(* IEC 61131-3 sources: plc-st-coding-agent/progress/evidence/f14_p1_20261111b/jobs/codex_minimax-m27 (part 2) *)

(* ---- public-easy-04.candidate_02.st ---- *)
PROGRAM JamPumpControl
VAR
    ViscosityDebounceTimer : TON;
    ViscosityConditionValid : BOOL := FALSE;
    FirstScan : BOOL := TRUE;
END_VAR

// Power-up initialization
IF FirstScan THEN
    VFD_RUN := FALSE;
    PUMP_RUNTIME_ACC := LTIME#0s;
    PUMP_MAINT_DUE := FALSE;
    ViscosityConditionValid := FALSE;
    FirstScan := FALSE;
END_IF;

// Viscosity debouncing logic
IF NOT VISCOSITY_OK THEN
    ViscosityConditionValid := FALSE;
    ViscosityDebounceTimer(IN := FALSE);
ELSE
    ViscosityDebounceTimer(IN := TRUE, PT := DebounceTime);
    IF ViscosityDebounceTimer.Q THEN
        ViscosityConditionValid := TRUE;
    END_IF;
END_IF;

// VFD_RUN control with E-STOP and viscosity permission
IF PASTE_E_STOP_NC AND ViscosityConditionValid THEN
    VFD_RUN := TRUE;
ELSE
    VFD_RUN := FALSE;
END_IF;

// Runtime accumulation while pump is running
IF VFD_RUN THEN
    PUMP_RUNTIME_ACC := PUMP_RUNTIME_ACC + CycleTime;
END_IF;

// Maintenance due indication at 500 hours
PUMP_MAINT_DUE := (PUMP_RUNTIME_ACC >= LTIME#500h);

END_PROGRAM

(* ---- public-easy-06.candidate_01.st ---- *)
PROGRAM AerationBlower
VAR
    // Inputs
    DO_LOW               : BOOL;  // Dissolved oxygen below threshold
    AERATION_E_STOP_NC   : BOOL;  // TRUE = E-stop inactive, FALSE = E-stop active

    // Outputs
    BLOWER_RUN                     : BOOL;  // Blower motor run command
    AERATION_BLOWER_CYCLE_COUNT    : UINT;  // Count of actual blower starts

    // Internal variables
    start_timer        : TON;      // On-delay timer for 5-second start delay
    blower_was_running : BOOL;     // Previous cycle state for edge detection
END_VAR

// Start delay: timer runs while both conditions are met
start_timer(
    IN := DO_LOW AND AERATION_E_STOP_NC,
    PT := T#5S
);

// Blower runs only when timer elapsed AND conditions remain satisfied
BLOWER_RUN := start_timer.Q AND DO_LOW AND AERATION_E_STOP_NC;

// Count FALSE-to-TRUE transitions of BLOWER_RUN (rising edge)
IF BLOWER_RUN AND NOT blower_was_running THEN
    AERATION_BLOWER_CYCLE_COUNT := AERATION_BLOWER_CYCLE_COUNT + 1;
END_IF;

// Update edge-detection state for next scan
blower_was_running := BLOWER_RUN;

END_PROGRAM

(* ---- public-hard-01.candidate_01.st ---- *)
// Material Proportioning Process Control - ST Implementation
// Supports Manual and Automatic modes with Emergency Stop

// ============================================================================
// Variable Declarations
// ============================================================================
VAR
    // System Inputs
    estop            : BOOL;   // Emergency Stop Signal (FALSE = triggered)
    opeMode          : BOOL;   // Operation Mode (FALSE = Manual, TRUE = Auto)
    valveAStart      : BOOL;   // Valve A Start Button
    valveBStart      : BOOL;   // Valve B Start Button
    valveCStart      : BOOL;   // Valve C Start Button
    valveDStart      : BOOL;   // Valve D Start Button
    mixMotorStart    : BOOL;   // Mixing Motor Start Button
    autoStart        : BOOL;   // Automatic Start Button
    processMode      : BOOL;   // Process Mode (FALSE = Basic, TRUE = Extended)
    levelSensor      : INT;    // Liquid Level Sensor (unit: cm)
    mixMotorComplete : BOOL;   // Mixing Complete Signal

    // System Outputs
    valveARun  : BOOL;   // Valve A Run Command
    valveBRun  : BOOL;   // Valve B Run Command
    valveCRun  : BOOL;   // Valve C Run Command
    valveDRun  : BOOL;   // Valve D Run Command
    mixMotorRun: BOOL;   // Mixing Motor Run Command

    // Internal Variables
    prevValveAStart   : BOOL;   // Previous state for edge detection
    prevValveBStart   : BOOL;
    prevValveCStart   : BOOL;
    prevValveDStart   : BOOL;
    prevMixMotorStart : BOOL;
    prevAutoStart     : BOOL;

    // Automatic Mode State Machine
    autoState : INT;     // 0=IDLE, 1=FILL_A, 2=FILL_B, 3=MIX_BASIC,
                         // 4=FILL_C, 5=MIX_EXT, 6=DRAIN
END_VAR

// ============================================================================
// Constants for State Machine
// ============================================================================
VAR CONSTANT
    STATE_IDLE      : INT := 0;
    STATE_FILL_A    : INT := 1;
    STATE_FILL_B    : INT := 2;
    STATE_MIX_BASIC : INT := 3;
    STATE_FILL_C    : INT := 4;
    STATE_MIX_EXT   : INT := 5;
    STATE_DRAIN     : INT := 6;
END_VAR

// ============================================================================
// Main Control Logic
// ============================================================================

// ---------------------------------------------------------------------------
// Emergency Stop Logic
// When estop=FALSE, all equipment stops immediately
// ---------------------------------------------------------------------------
IF NOT estop THEN
    // Emergency stop: immediate shutdown of all outputs
    valveARun  := FALSE;
    valveBRun  := FALSE;
    valveCRun  := FALSE;
    valveDRun  := FALSE;
    mixMotorRun:= FALSE;
    autoState  := STATE_IDLE;

    // Reset edge detection flags to prevent spurious triggers after estop release
    prevValveAStart   := FALSE;
    prevValveBStart   := FALSE;
    prevValveCStart   := FALSE;
    prevValveDStart   := FALSE;
    prevMixMotorStart := FALSE;
    prevAutoStart     := FALSE;
    RETURN;  // Skip remaining logic when emergency stop is active
END_IF

// ---------------------------------------------------------------------------
// Mode Selection: Manual vs Automatic
// ---------------------------------------------------------------------------
IF NOT opeMode THEN
    // ============================
    // MANUAL OPERATION MODE
    // Toggle each device on rising edge of corresponding button
    // ============================

    // Valve A Toggle Control
    IF valveAStart AND NOT prevValveAStart THEN
        valveARun := NOT valveARun;
    END_IF
    prevValveAStart := valveAStart;

    // Valve B Toggle Control
    IF valveBStart AND NOT prevValveBStart THEN
        valveBRun := NOT valveBRun;
    END_IF
    prevValveBStart := valveBStart;

    // Valve C Toggle Control
    IF valveCStart AND NOT prevValveCStart THEN
        valveCRun := NOT valveCRun;
    END_IF
    prevValveCStart := valveCStart;

    // Valve D Toggle Control
    IF valveDStart AND NOT prevValveDStart THEN
        valveDRun := NOT valveDRun;
    END_IF
    prevValveDStart := valveDStart;

    // Mixing Motor Toggle Control
    IF mixMotorStart AND NOT prevMixMotorStart THEN
        mixMotorRun := NOT mixMotorRun;
    END_IF
    prevMixMotorStart := mixMotorStart;

ELSE
    // ============================
    // AUTOMATIC OPERATION MODE
    // Sequential process control based on state machine
    // ============================

    // Reset manual control outputs when switching to auto mode
    valveARun  := FALSE;
    valveBRun  := FALSE;
    valveCRun  := FALSE;
    valveDRun  := FALSE;
    mixMotorRun:= FALSE;

    // Start automatic process on rising edge of autoStart button
    IF autoStart AND NOT prevAutoStart THEN
        IF autoState = STATE_IDLE THEN
            autoState := STATE_FILL_A;  // Begin the automatic sequence
        END_IF
    END_IF
    prevAutoStart := autoStart;

    // ---------------------------------------------------------------------------
    // Automatic Mode State Machine
    // ---------------------------------------------------------------------------
    CASE autoState OF

        STATE_IDLE:
            // Wait for autoStart button press
            valveARun  := FALSE;
            valveBRun  := FALSE;
            valveCRun  := FALSE;
            valveDRun  := FALSE;
            mixMotorRun:= FALSE;

        STATE_FILL_A:
            // Open Valve A to fill tank
            valveARun := TRUE;
            valveBRun := FALSE;
            valveCRun := FALSE;
            valveDRun := FALSE;
            mixMotorRun := FALSE;

            // When level reaches 50cm, close Valve A and proceed to Valve B
            IF levelSensor >= 50 THEN
                valveARun := FALSE;
                autoState := STATE_FILL_B;
            END_IF

        STATE_FILL_B:
            // Open Valve B to continue filling
            valveARun := FALSE;
            valveBRun := TRUE;
            valveCRun := FALSE;
            valveDRun := FALSE;
            mixMotorRun := FALSE;

            // When level reaches 80cm, close Valve B
            IF levelSensor >= 80 THEN
                valveBRun := FALSE;

                // Branch based on processMode
                IF NOT processMode THEN
                    // Basic Mode: Start mixing directly
                    autoState := STATE_MIX_BASIC;
                ELSE
                    // Extended Mode: Open Valve C for additional fill
                    autoState := STATE_FILL_C;
                END_IF
            END_IF

        STATE_MIX_BASIC:
            // Basic Mode: Start mixing motor
            valveARun  := FALSE;
            valveBRun  := FALSE;
            valveCRun  := FALSE;
            valveDRun  := FALSE;
            mixMotorRun := TRUE;

            // When mixing complete, stop motor and open drain valve
            IF mixMotorComplete THEN
                mixMotorRun := FALSE;
                autoState := STATE_DRAIN;
            END_IF

        STATE_FILL_C:
            // Extended Mode: Open Valve C for additional material
            valveARun  := FALSE;
            valveBRun  := FALSE;
            valveCRun  := TRUE;
            valveDRun  := FALSE;
            mixMotorRun := FALSE;

            // When level reaches 100cm, close Valve C and start mixing
            IF levelSensor >= 100 THEN
                valveCRun := FALSE;
                autoState := STATE_MIX_EXT;
            END_IF

        STATE_MIX_EXT:
            // Extended Mode: Start mixing motor
            valveARun  := FALSE;
            valveBRun  := FALSE;
            valveCRun  := FALSE;
            valveDRun  := FALSE;
            mixMotorRun := TRUE;

            // When mixing complete, stop motor and open drain valve
            IF mixMotorComplete THEN
                mixMotorRun := FALSE;
                autoState := STATE_DRAIN;
            END_IF

        STATE_DRAIN:
            // Open Valve D to drain tank (deliver to next process)
            valveARun  := FALSE;
            valveBRun  := FALSE;
            valveCRun  := FALSE;
            valveDRun  := TRUE;
            mixMotorRun := FALSE;

            // Return to idle when tank is empty (level < 10cm)
            IF levelSensor < 10 THEN
                valveDRun := FALSE;
                autoState := STATE_IDLE;  // Process complete, ready for next cycle
            END_IF

    END_CASE

END_IF

(* ---- public-hard-02.candidate_01.st ---- *)
I'll implement the Flexible Processing Control system in Structured Text (ST). Let me analyze the requirements and create a complete solution.

## Analysis

This is a state-machine-based conveyor control system with:
- 5 stations (1# loading, 2#-4# processing, 5# output)
- Event-driven transitions based on sensors and completion signals
- Process sequence control from input array
- Direction control for conveyor movement

I'll create a complete ST program with proper state management and edge-triggered logic to prevent multiple activations.
<file_write file="FlexibleProcessingControl.st">
PROGRAM FlexibleProcessingControl
VAR
    // Inputs
    processLength     : USINT;                      // Active process-sequence length, 1..8
    sensor1, sensor2, sensor3, sensor4, sensor5 : BOOL;  // Station sensors
    station1Start     : BOOL;                       // Start button at 1# station
    station2Complete  : BOOL;                       // Processing completion at 2#
    station3Complete  : BOOL;                       // Processing completion at 3#
    station4Complete  : BOOL;                       // Processing completion at 4#
    processSequence   : ARRAY[1..8] OF USINT;       // Processing sequence array

    // Outputs
    conveyorLeft      : BOOL;                       // Conveyor moves left
    conveyorRight     : BOOL;                       // Conveyor moves right

    // Internal variables
    currentStep       : USINT := 1;                 // Current step in process sequence
    currentPosition   : USINT := 1;                 // Current station position (1-5)
    isRunning         : BOOL := FALSE;              // Processing state flag
    targetStation     : USINT;                      // Target station for current move

    // Edge detection flags for completion signals
    station2CompletePrev : BOOL := FALSE;
    station3CompletePrev : BOOL := FALSE;
    station4CompletePrev : BOOL := FALSE;

    // State machine states
    STATE_IDLE        : USINT := 0;
    STATE_MOVING      : USINT := 1;
    STATE_WAITING     : USINT := 2;
    currentState      : USINT := STATE_IDLE;
END_VAR

// ============================================================================
// Main Control Logic
// ============================================================================

// --------------------------------------------------------------------
// State: IDLE
// Wait for start button at station 1 with raw material detected
// --------------------------------------------------------------------
IF currentState = STATE_IDLE THEN
    // Check if start button is pressed with material at station 1
    IF sensor1 AND station1Start AND NOT isRunning THEN
        // Initialize process
        isRunning := TRUE;
        currentStep := 1;
        currentPosition := 1;

        // Check if process sequence is valid
        IF processLength >= 1 AND processLength <= 8 THEN
            // Get first target from process sequence
            targetStation := processSequence[currentStep];

            // Validate target station (should be 2-5)
            IF targetStation >= 2 AND targetStation <= 5 THEN
                currentState := STATE_MOVING;
            ELSE
                // Invalid sequence, abort
                isRunning := FALSE;
                currentState := STATE_IDLE;
            END_IF
        ELSE
            // Invalid process length, abort
            isRunning := FALSE;
            currentState := STATE_IDLE;
        END_IF
    END_IF

// --------------------------------------------------------------------
// State: MOVING
// Control conveyor direction to move product to target station
// --------------------------------------------------------------------
ELSIF currentState = STATE_MOVING THEN
    // Determine conveyor direction based on target station
    IF targetStation > currentPosition THEN
        // Need to move right (forward)
        conveyorRight := TRUE;
        conveyorLeft := FALSE;
    ELSIF targetStation < currentPosition THEN
        // Need to move left (backward)
        conveyorLeft := TRUE;
        conveyorRight := FALSE;
    ELSE
        // Already at target, stop conveyor
        conveyorLeft := FALSE;
        conveyorRight := FALSE;
        currentState := STATE_WAITING;
    END_IF

// --------------------------------------------------------------------
// State: WAITING
// Wait for product to arrive at target station
// Then wait for processing completion (for stations 2-4)
// --------------------------------------------------------------------
ELSIF currentState = STATE_WAITING THEN
    // Stop conveyor while waiting
    conveyorLeft := FALSE;
    conveyorRight := FALSE;

    // Check product arrival at target station
    IF (targetStation = 2 AND sensor2) OR
       (targetStation = 3 AND sensor3) OR
       (targetStation = 4 AND sensor4) OR
       (targetStation = 5 AND sensor5) THEN
        // Product has arrived at target station
        currentPosition := targetStation;

        // Check if this is the final station (5#)
        IF targetStation = 5 THEN
            // Process complete - reset to idle
            isRunning := FALSE;
            currentStep := 1;
            currentState := STATE_IDLE;
        ELSE
            // For stations 2-4, wait for completion signal
            // State remains WAITING until completion signal received
        END_IF
    END_IF
END_IF

// ============================================================================
// Process Completion Handling (checked in every state)
// ============================================================================

// Handle station 2 completion with edge detection
IF station2Complete AND NOT station2CompletePrev THEN
    IF isRunning AND currentPosition = 2 THEN
        // Station 2 completed, advance to next step
        currentStep := currentStep + 1;

        // Check if process is complete
        IF currentStep > processLength THEN
            // Should not happen if sequence ends at station 5
            isRunning := FALSE;
            currentStep := 1;
            currentState := STATE_IDLE;
        ELSE
            // Get next target from process sequence
            targetStation := processSequence[currentStep];

            // Validate target station
            IF targetStation >= 2 AND targetStation <= 5 THEN
                currentState := STATE_MOVING;
            ELSE
                // Invalid sequence, abort
                isRunning := FALSE;
                currentStep := 1;
                currentState := STATE_IDLE;
            END_IF
        END_IF
    END_IF
END_IF
station2CompletePrev := station2Complete;

// Handle station 3 completion with edge detection
IF station3Complete AND NOT station3CompletePrev THEN
    IF isRunning AND currentPosition = 3 THEN
        // Station 3 completed, advance to next step
        currentStep := currentStep + 1;

        // Check if process is complete
        IF currentStep > processLength THEN
            // Should not happen if sequence ends at station 5
            isRunning := FALSE;
            currentStep := 1;
            currentState := STATE_IDLE;
        ELSE
            // Get next target from process sequence
            targetStation := processSequence[currentStep];

            // Validate target station
            IF targetStation >= 2 AND targetStation <= 5 THEN
                currentState := STATE_MOVING;
            ELSE
                // Invalid sequence, abort
                isRunning := FALSE;
                currentStep := 1;
                currentState := STATE_IDLE;
            END_IF
        END_IF
    END_IF
END_IF
station3CompletePrev := station3Complete;

// Handle station 4 completion with edge detection
IF station4Complete AND NOT station4CompletePrev THEN
    IF isRunning AND currentPosition = 4 THEN
        // Station 4 completed, advance to next step
        currentStep := currentStep + 1;

        // Check if process is complete
        IF currentStep > processLength THEN
            // Should not happen if sequence ends at station 5
            isRunning := FALSE;
            currentStep := 1;
            currentState := STATE_IDLE;
        ELSE
            // Get next target from process sequence
            targetStation := processSequence[currentStep];

            // Validate target station
            IF targetStation >= 2 AND targetStation <= 5 THEN
                currentState := STATE_MOVING;
            ELSE
                // Invalid sequence, abort
                isRunning := FALSE;
                currentStep := 1;
                currentState := STATE_IDLE;
            END_IF
        END_IF
    END_IF
END_IF
station4CompletePrev := station4Complete;

END_PROGRAM
</file_write>

**Key implementation details:**

1. **State Machine** with three states:
   - `STATE_IDLE`: Waiting for start button with material at station 1
   - `STATE_MOVING`: Conveyor active, moving to target station
   - `STATE_WAITING`: Product at station, waiting for completion signal (2-4) or completion (5)

2. **Edge-triggered completion signals** using `_Prev` flags to prevent multiple activations

3. **Conveyor direction logic**: Compares `targetStation` vs `currentPosition` to determine left/right movement

4. **Process sequence validation**: Ensures target stations are in valid range (2-5)

5. **Auto-reset**: When product reaches station 5, system returns to idle state and is ready for next product

The program assumes that once the product reaches station 5 (output), the external system removes it, causing `sensor5` to go false, making the system ready for the next product.

(* ---- public-hard-02.candidate_02.st ---- *)
I'll fix the backtick characters that aren't valid in ST and provide the corrected code.
<file_write file="FlexibleProcessingControl.st">
PROGRAM FlexibleProcessingControl
VAR
    processLength     : USINT;
    sensor1, sensor2, sensor3, sensor4, sensor5 : BOOL;
    station1Start     : BOOL;
    station2Complete  : BOOL;
    station3Complete  : BOOL;
    station4Complete  : BOOL;
    processSequence   : ARRAY[1..8] OF USINT;

    conveyorLeft      : BOOL;
    conveyorRight     : BOOL;

    currentStep       : USINT := 1;
    currentPosition   : USINT := 1;
    isRunning         : BOOL := FALSE;
    targetStation     : USINT;

    station2CompletePrev : BOOL := FALSE;
    station3CompletePrev : BOOL := FALSE;
    station4CompletePrev : BOOL := FALSE;

    STATE_IDLE        : USINT := 0;
    STATE_MOVING      : USINT := 1;
    STATE_WAITING     : USINT := 2;
    currentState      : USINT := 0;
END_VAR

IF currentState = STATE_IDLE THEN
    IF sensor1 AND station1Start AND NOT isRunning THEN
        isRunning := TRUE;
        currentStep := 1;
        currentPosition := 1;

        IF processLength >= 1 AND processLength <= 8 THEN
            targetStation := processSequence[currentStep];

            IF targetStation >= 2 AND targetStation <= 5 THEN
                currentState := STATE_MOVING;
            ELSE
                isRunning := FALSE;
                currentState := STATE_IDLE;
            END_IF
        ELSE
            isRunning := FALSE;
            currentState := STATE_IDLE;
        END_IF
    END_IF

ELSIF currentState = STATE_MOVING THEN
    IF targetStation > currentPosition THEN
        conveyorRight := TRUE;
        conveyorLeft := FALSE;
    ELSIF targetStation < currentPosition THEN
        conveyorLeft := TRUE;
        conveyorRight := FALSE;
    ELSE
        conveyorLeft := FALSE;
        conveyorRight := FALSE;
        currentState := STATE_WAITING;
    END_IF

ELSIF currentState = STATE_WAITING THEN
    conveyorLeft := FALSE;
    conveyorRight := FALSE;

    IF (targetStation = 2 AND sensor2) OR
       (targetStation = 3 AND sensor3) OR
       (targetStation = 4 AND sensor4) OR
       (targetStation = 5 AND sensor5) THEN
        currentPosition := targetStation;

        IF targetStation = 5 THEN
            isRunning := FALSE;
            currentStep := 1;
            currentState := STATE_IDLE;
        END_IF
    END_IF
END_IF

IF station2Complete AND NOT station2CompletePrev THEN
    IF isRunning AND currentPosition = 2 THEN
        currentStep := currentStep + 1;

        IF currentStep > processLength THEN
            isRunning := FALSE;
            currentStep := 1;
            currentState := STATE_IDLE;
        ELSE
            targetStation := processSequence[currentStep];

            IF targetStation >= 2 AND targetStation <= 5 THEN
                currentState := STATE_MOVING;
            ELSE
                isRunning := FALSE;
                currentStep := 1;
                currentState := STATE_IDLE;
            END_IF
        END_IF
    END_IF
END_IF
station2CompletePrev := station2Complete;

IF station3Complete AND NOT station3CompletePrev THEN
    IF isRunning AND currentPosition = 3 THEN
        currentStep := currentStep + 1;

        IF currentStep > processLength THEN
            isRunning := FALSE;
            currentStep := 1;
            currentState := STATE_IDLE;
        ELSE
            targetStation := processSequence[currentStep];

            IF targetStation >= 2 AND targetStation <= 5 THEN
                currentState := STATE_MOVING;
            ELSE
                isRunning := FALSE;
                currentStep := 1;
                currentState := STATE_IDLE;
            END_IF
        END_IF
    END_IF
END_IF
station3CompletePrev := station3Complete;

IF station4Complete AND NOT station4CompletePrev THEN
    IF isRunning AND currentPosition = 4 THEN
        currentStep := currentStep + 1;

        IF currentStep > processLength THEN
            isRunning := FALSE;
            currentStep := 1;
            currentState := STATE_IDLE;
        ELSE
            targetStation := processSequence[currentStep];

            IF targetStation >= 2 AND targetStation <= 5 THEN
                currentState := STATE_MOVING;
            ELSE
                isRunning := FALSE;
                currentStep := 1;
                currentState := STATE_IDLE;
            END_IF
        END_IF
    END_IF
END_IF
station4CompletePrev := station4Complete;

END_PROGRAM
</file_write>

(* ---- public-hard-03.candidate_01.st ---- *)
PROGRAM RecipeManagement
VAR
    // Inputs
    addRecipe     : BOOL;
    deleteRecipe  : BOOL;
    modifyRecipe  : BOOL;
    queryRecipe   : BOOL;
    recipeIn      : ST_Recipe;

    // Outputs
    recipeAdded         : BOOL;
    recipeDeleted       : BOOL;
    recipeModified      : BOOL;
    recipeQueryResult   : ST_Recipe;
    error               : BOOL;
    status              : WORD;

    // Internal variables
    recipe              : ARRAY[1..10] OF ST_Recipe;
    i                   : INT;
    foundIndex          : INT;
    emptySlotIndex      : INT;
END_VAR
// Implementation
// Initialize internal tracking variables
foundIndex := 0;
emptySlotIndex := 0;

// Reset all output signals
recipeAdded := FALSE;
recipeDeleted := FALSE;
recipeModified := FALSE;
error := FALSE;
status := 16#0000;

// Search for existing recipe and find first empty slot
FOR i := 1 TO 10 DO
    IF recipe[i].recipeID <> 0 THEN
        // This slot contains a recipe
        IF recipe[i].recipeID = recipeIn.recipeID THEN
            foundIndex := i;
        END_IF
    ELSE
        // This is an empty slot
        IF emptySlotIndex = 0 THEN
            emptySlotIndex := i;
        END_IF
    END_IF
END_FOR;

// Handle Query Recipe Request
IF queryRecipe THEN
    IF foundIndex <> 0 THEN
        // Recipe found - output it
        recipeQueryResult := recipe[foundIndex];
    ELSE
        // Recipe not found - error
        error := TRUE;
        status := 16#8001;
    END_IF
END_IF

// Handle Add Recipe Request
IF addRecipe THEN
    IF foundIndex <> 0 THEN
        // Duplicate recipe number found - error
        error := TRUE;
        status := 16#8002;
    ELSIF emptySlotIndex = 0 THEN
        // No empty slot available - error
        error := TRUE;
        status := 16#8003;
    ELSE
        // Add recipe to the first empty slot
        recipe[emptySlotIndex] := recipeIn;
        recipeAdded := TRUE;
    END_IF
END_IF

// Handle Delete Recipe Request
IF deleteRecipe THEN
    IF foundIndex <> 0 THEN
        // Recipe found - delete it by setting recipeID to 0
        recipe[foundIndex].recipeID := 0;
        recipeDeleted := TRUE;
    ELSE
        // Recipe not found - error
        error := TRUE;
        status := 16#8004;
    END_IF
END_IF

// Handle Modify Recipe Request
IF modifyRecipe THEN
    IF foundIndex <> 0 THEN
        // Recipe found - replace with input recipe
        recipe[foundIndex] := recipeIn;
        recipeModified := TRUE;
    ELSE
        // Recipe not found - error
        error := TRUE;
        status := 16#8005;
    END_IF
END_IF

(* ---- public-hard-03.candidate_02.st ---- *)
PROGRAM RecipeManagement
VAR
    // Inputs
    addRecipe     : BOOL;
    deleteRecipe  : BOOL;
    modifyRecipe  : BOOL;
    queryRecipe   : BOOL;
    recipeIn      : ST_Recipe;

    // Outputs
    recipeAdded         : BOOL;
    recipeDeleted       : BOOL;
    recipeModified      : BOOL;
    recipeQueryResult   : ST_Recipe;
    error               : BOOL;
    status              : WORD;

    // Internal variables
    recipe              : ARRAY[1..10] OF ST_Recipe;
    i                   : INT;
    foundIndex          : INT;
    emptySlotIndex      : INT;
END_VAR
// Implementation
// Initialize internal tracking variables
foundIndex := 0;
emptySlotIndex := 0;

// Reset all output signals
recipeAdded := FALSE;
recipeDeleted := FALSE;
recipeModified := FALSE;
error := FALSE;
status := 16#0000;

// Search for existing recipe and find first empty slot
FOR i := 1 TO 10 DO
    IF recipe[i].recipeID <> 0 THEN
        // This slot contains a recipe
        IF recipe[i].recipeID = recipeIn.recipeID THEN
            foundIndex := i;
        END_IF
    ELSE
        // This is an empty slot
        IF emptySlotIndex = 0 THEN
            emptySlotIndex := i;
        END_IF
    END_IF
END_FOR;

// Handle Query Recipe Request
IF queryRecipe THEN
    IF foundIndex <> 0 THEN
        // Recipe found - output it
        recipeQueryResult := recipe[foundIndex];
    ELSE
        // Recipe not found - error
        error := TRUE;
        status := 16#8001;
    END_IF
END_IF

// Handle Add Recipe Request
IF addRecipe THEN
    IF foundIndex <> 0 THEN
        // Duplicate recipe number found - error
        error := TRUE;
        status := 16#8002;
    ELSIF emptySlotIndex = 0 THEN
        // No empty slot available - error
        error := TRUE;
        status := 16#8003;
    ELSE
        // Add recipe to the first empty slot
        recipe[emptySlotIndex] := recipeIn;
        recipeAdded := TRUE;
    END_IF
END_IF

// Handle Delete Recipe Request
IF deleteRecipe THEN
    IF foundIndex <> 0 THEN
        // Recipe found - delete it by setting recipeID to 0
        recipe[foundIndex].recipeID := 0;
        recipeDeleted := TRUE;
    ELSE
        // Recipe not found - error
        error := TRUE;
        status := 16#8004;
    END_IF
END_IF

// Handle Modify Recipe Request
IF modifyRecipe THEN
    IF foundIndex <> 0 THEN
        // Recipe found - replace with input recipe
        recipe[foundIndex] := recipeIn;
        recipeModified := TRUE;
    ELSE
        // Recipe not found - error
        error := TRUE;
        status := 16#8005;
    END_IF
END_IF

END_PROGRAM

(* ---- public-hard-04.candidate_01.st ---- *)
METHOD GetBufferInfo : BOOL
VAR_INPUT
    buffer : VARIANT;
END_VAR
VAR_OUTPUT
    capacity    : DINT;
    elementSize : DINT;
END_VAR

VAR
    pBuffer    : REFERENCE TO BYTE;
    bufferType : REF_TO ANY;
END_VAR

bufferType REF= buffer;

IF __ISVALIDREF(bufferType) THEN
    capacity := bufferType.GetUpperBound(1) + 1;
    elementSize := bufferType.GetSize() / capacity;
    GetBufferInfo := TRUE;
ELSE
    capacity := 0;
    elementSize := 0;
    GetBufferInfo := FALSE;
END_IF
END_METHOD

METHOD Enqueue : BOOL
VAR_INPUT
    buffer      : VARIANT;
    item        : VARIANT;
    tail        : DINT;
    elementCount: DINT;
    elementSize : DINT;
END_VAR

VAR
    pDest : POINTER TO BYTE;
    pSrc  : POINTER TO BYTE;
    idx   : DINT;
END_VAR

idx := tail MOD THIS^._capacity;

pDest := __GET_VAR_DATA_REF(buffer).ADR + (idx * elementSize);
pSrc  := __GET_VAR_DATA_REF(item).ADR;

MemMove(pSrc, pDest, elementSize);

THIS^._tail := (tail + 1) MOD THIS^._capacity;
THIS^._elementCount := elementCount + 1;

Enqueue := TRUE;
END_METHOD

METHOD Dequeue : BOOL
VAR_INPUT
    buffer      : VARIANT;
    item        : VARIANT;
    head        : DINT;
    elementCount: DINT;
    elementSize : DINT;
END_VAR

VAR
    pSrc  : POINTER TO BYTE;
    pDest : POINTER TO BYTE;
    idx   : DINT;
    zeroBuf : ARRAY[0..255] OF BYTE;
END_VAR

idx := head MOD THIS^._capacity;

pSrc  := __GET_VAR_DATA_REF(buffer).ADR + (idx * elementSize);
pDest := __GET_VAR_DATA_REF(item).ADR;

MemMove(pSrc, pDest, elementSize);

MemSet(zeroBuf, 0, elementSize);
MemMove(zeroBuf, pSrc, elementSize);

THIS^._head := (head + 1) MOD THIS^._capacity;
THIS^._elementCount := elementCount - 1;

Dequeue := TRUE;
END_METHOD

(* ---- public-hard-06.candidate_01.st ---- *)
(* Production Line Control System *)
(* 5 Workstations: Loading → Cleaning → Weighing → Firing → Finished Product *)

PROGRAM ProductionLineControl
VAR
    (* Mode Selection *)
    Mode AT %IX0.0 : BOOL;              (* 0=Manual, 1=Automatic *)

    (* Manual Mode Inputs *)
    ForwardButton AT %IX0.1 : BOOL;     (* Forward rotation button *)
    ReverseButton AT %IX0.2 : BOOL;     (* Reverse rotation button *)

    (* Automatic Mode - Sensors *)
    SensorFeed AT %IX0.3 : BOOL;        (* Material loading station sensor *)
    SensorWash AT %IX0.4 : BOOL;        (* Cleaning station sensor *)
    SensorWeight AT %IX0.5 : BOOL;      (* Weighing station sensor *)
    SensorFiring AT %IX0.6 : BOOL;      (* Firing station sensor *)
    SensorOutput AT %IX0.7 : BOOL;      (* Finished product station sensor *)

    (* Process Completion Signals *)
    washComplete AT %IX1.0 : BOOL;      (* Cleaning complete signal *)
    weightComplete AT %IX1.1 : BOOL;    (* Weighing complete signal *)
    firingComplete AT %IX1.2 : BOOL;    (* Firing complete signal *)

    (* Process Values *)
    weight AT %ID2 : REAL;              (* Weight value (REAL type) *)

    (* Outputs *)
    MotorForward AT %QX0.0 : BOOL;      (* Motor forward rotation *)
    MotorReverse AT %QX0.1 : BOOL;      (* Motor reverse rotation *)
    kick AT %QX0.2 : BOOL;              (* Rejection output *)
    CompletionLight AT %QX0.3 : BOOL;   (* Completion indicator light *)
    firingTemp AT %QD2 : REAL;          (* Firing temperature (REAL type) *)

    (* State Machine Variables *)
    CurrentState : INT;
    PreviousSensorFeed : BOOL;
    PreviousSensorWash : BOOL;
    PreviousSensorWeight : BOOL;
    PreviousSensorFiring : BOOL;
    PreviousSensorOutput : BOOL;
    PreviousWashComplete : BOOL;
    PreviousWeightComplete : BOOL;
    PreviousFiringComplete : BOOL;

    (* Edge Detection Flags *)
    SensorFeedEdge : BOOL;
    SensorWashEdge : BOOL;
    SensorWeightEdge : BOOL;
    SensorFiringEdge : BOOL;
    SensorOutputEdge : BOOL;
    WashCompleteEdge : BOOL;
    WeightCompleteEdge : BOOL;
    FiringCompleteEdge : BOOL;

    (* Temporary Variables *)
    weightValue : REAL;
    tempCalc : REAL;
END_VAR

(* Constants for States *)
CONST
    STATE_IDLE : INT := 0;
    STATE_FEED_DETECTED : INT := 1;
    STATE_WASH_WAIT : INT := 2;
    STATE_WEIGHING_WAIT : INT := 3;
    STATE_WEIGHT_CHECK : INT := 4;
    STATE_FIRING_WAIT : INT := 5;
    STATE_OUTPUT_WAIT : INT := 6;
END_CONST

(* Main Control Logic *)
(* -------------------------------------------------------- *)
(* EDGE DETECTION FOR ALL SENSORS AND SIGNALS *)
SensorFeedEdge := SensorFeed AND NOT PreviousSensorFeed;
SensorWashEdge := SensorWash AND NOT PreviousSensorWash;
SensorWeightEdge := SensorWeight AND NOT PreviousSensorWeight;
SensorFiringEdge := SensorFiring AND NOT PreviousSensorFiring;
SensorOutputEdge := SensorOutput AND NOT PreviousSensorOutput;
WashCompleteEdge := washComplete AND NOT PreviousWashComplete;
WeightCompleteEdge := weightComplete AND NOT PreviousWeightComplete;
FiringCompleteEdge := firingComplete AND NOT PreviousFiringComplete;

(* Update Previous States *)
PreviousSensorFeed := SensorFeed;
PreviousSensorWash := SensorWash;
PreviousSensorWeight := SensorWeight;
PreviousSensorFiring := SensorFiring;
PreviousSensorOutput := SensorOutput;
PreviousWashComplete := washComplete;
PreviousWeightComplete := weightComplete;
PreviousFiringComplete := firingComplete;

(* -------------------------------------------------------- *)
(* MANUAL MODE CONTROL *)
IF Mode = FALSE THEN
    (* Interlock: Forward and Reverse cannot be active simultaneously *)
    MotorForward := ForwardButton AND NOT ReverseButton;
    MotorReverse := ReverseButton AND NOT ForwardButton;

    (* Reset automatic mode outputs *)
    kick := FALSE;
    CompletionLight := FALSE;
    firingTemp := 0.0;

    (* Reset state machine *)
    CurrentState := STATE_IDLE;
END_IF

(* -------------------------------------------------------- *)
(* AUTOMATIC MODE CONTROL *)
IF Mode = TRUE THEN
    CASE CurrentState OF

        (* STATE_IDLE: Wait for material at loading station *)
        STATE_IDLE:
            MotorForward := FALSE;
            MotorReverse := FALSE;
            kick := FALSE;
            CompletionLight := FALSE;
            firingTemp := 0.0;

            (* Material detected at loading station *)
            IF SensorFeedEdge THEN
                CurrentState := STATE_FEED_DETECTED;
            END_IF

        (* STATE_FEED_DETECTED: Material detected, start motor to move to cleaning *)
        STATE_FEED_DETECTED:
            MotorForward := TRUE;
            MotorReverse := FALSE;
            kick := FALSE;
            CompletionLight := FALSE;

            (* Material reached cleaning station *)
            IF SensorWashEdge THEN
                MotorForward := FALSE;
                CurrentState := STATE_WASH_WAIT;
            END_IF

        (* STATE_WASH_WAIT: Material at cleaning station, wait for washComplete *)
        STATE_WASH_WAIT:
            MotorForward := FALSE;
            MotorReverse := FALSE;
            kick := FALSE;
            CompletionLight := FALSE;

            (* Cleaning complete, move to weighing *)
            IF WashCompleteEdge THEN
                MotorForward := TRUE;
                CurrentState := STATE_WEIGHING_WAIT;
            END_IF

        (* STATE_WEIGHING_WAIT: Material at weighing station, wait for weightComplete *)
        STATE_WEIGHING_WAIT:
            MotorForward := FALSE;
            MotorReverse := FALSE;
            kick := FALSE;
            CompletionLight := FALSE;

            (* Weighing complete, check weight *)
            IF WeightCompleteEdge THEN
                CurrentState := STATE_WEIGHT_CHECK;
            END_IF

        (* STATE_WEIGHT_CHECK: Evaluate weight and determine qualification *)
        STATE_WEIGHT_CHECK:
            weightValue := weight;

            (* Check if weight is within qualified range [100, 200] *)
            IF (weightValue >= 100.0) AND (weightValue <= 200.0) THEN
                (* Qualified product - Calculate firing temperature *)
                (* Linear mapping: weight 100→200 maps to temperature 500→550 *)
                tempCalc := 500.0 + ((weightValue - 100.0) / 100.0) * 50.0;
                firingTemp := tempCalc;
                kick := FALSE;

                (* Move to firing station *)
                MotorForward := TRUE;
                MotorReverse := FALSE;
                CurrentState := STATE_FIRING_WAIT;
            ELSE
                (* Unqualified product - Reject *)
                kick := TRUE;
                firingTemp := 0.0;
                MotorForward := FALSE;
                MotorReverse := FALSE;

                (* Return to idle after rejection *)
                CurrentState := STATE_IDLE;
            END_IF

        (* STATE_FIRING_WAIT: Product at firing station, wait for firingComplete *)
        STATE_FIRING_WAIT:
            kick := FALSE;
            CompletionLight := FALSE;

            (* Keep firing temperature active during firing *)
            IF firingTemp > 0.0 THEN
                (* Firing in progress, maintain temperature output *)
            END_IF;

            (* Firing complete, move to finished product station *)
            IF FiringCompleteEdge THEN
                MotorForward := TRUE;
                MotorReverse := FALSE;
                CurrentState := STATE_OUTPUT_WAIT;
            END_IF

        (* STATE_OUTPUT_WAIT: Product at finished product station *)
        STATE_OUTPUT_WAIT:
            MotorForward := FALSE;
            MotorReverse := FALSE;
            kick := FALSE;

            (* Product detected at output - Turn on completion light *)
            IF SensorOutput THEN
                CompletionLight := TRUE;
            ELSE
                (* Product taken away - Turn off completion light *)
                CompletionLight := FALSE;
                CurrentState := STATE_IDLE;
            END_IF

    END_CASE
END_IF

(* -------------------------------------------------------- *)
(* SAFETY: Emergency Stop Logic - Disable outputs if in error state *)
(* (This can be extended based on additional safety requirements) *)

END_PROGRAM

(* ---- public-hard-06.candidate_02.st ---- *)
(* Production Line Control System *)
(* 5 Workstations: Loading → Cleaning → Weighing → Firing → Finished Product *)

PROGRAM ProductionLineControl
VAR
    (* Mode Selection *)
    Mode AT %IX0.0 : BOOL;              (* 0=Manual, 1=Automatic *)

    (* Manual Mode Inputs *)
    ForwardButton AT %IX0.1 : BOOL;     (* Forward rotation button *)
    ReverseButton AT %IX0.2 : BOOL;     (* Reverse rotation button *)

    (* Automatic Mode - Sensors *)
    SensorFeed AT %IX0.3 : BOOL;        (* Material loading station sensor *)
    SensorWash AT %IX0.4 : BOOL;        (* Cleaning station sensor *)
    SensorWeight AT %IX0.5 : BOOL;      (* Weighing station sensor *)
    SensorFiring AT %IX0.6 : BOOL;      (* Firing station sensor *)
    SensorOutput AT %IX0.7 : BOOL;      (* Finished product station sensor *)

    (* Process Completion Signals *)
    washComplete AT %IX1.0 : BOOL;      (* Cleaning complete signal *)
    weightComplete AT %IX1.1 : BOOL;    (* Weighing complete signal *)
    firingComplete AT %IX1.2 : BOOL;    (* Firing complete signal *)

    (* Process Values *)
    weight AT %ID2 : REAL;              (* Weight value *)

    (* Outputs *)
    MotorForward AT %QX0.0 : BOOL;      (* Motor forward rotation *)
    MotorReverse AT %QX0.1 : BOOL;      (* Motor reverse rotation *)
    kick AT %QX0.2 : BOOL;              (* Rejection output *)
    CompletionLight AT %QX0.3 : BOOL;   (* Completion indicator light *)
    firingTemp AT %QD2 : REAL;          (* Firing temperature *)

    (* State Machine Variables *)
    CurrentState : INT;
    PreviousSensorFeed : BOOL;
    PreviousSensorWash : BOOL;
    PreviousSensorWeight : BOOL;
    PreviousSensorFiring : BOOL;
    PreviousSensorOutput : BOOL;
    PreviousWashComplete : BOOL;
    PreviousWeightComplete : BOOL;
    PreviousFiringComplete : BOOL;

    (* Edge Detection Flags *)
    SensorFeedEdge : BOOL;
    SensorWashEdge : BOOL;
    SensorWeightEdge : BOOL;
    SensorFiringEdge : BOOL;
    SensorOutputEdge : BOOL;
    WashCompleteEdge : BOOL;
    WeightCompleteEdge : BOOL;
    FiringCompleteEdge : BOOL;

    (* Temporary Variables *)
    weightValue : REAL;
    tempCalc : REAL;
END_VAR

(* Constants for States *)
VAR CONSTANT
    STATE_IDLE : INT := 0;
    STATE_FEED_DETECTED : INT := 1;
    STATE_WASH_WAIT : INT := 2;
    STATE_WEIGHING_WAIT : INT := 3;
    STATE_WEIGHT_CHECK : INT := 4;
    STATE_FIRING_WAIT : INT := 5;
    STATE_OUTPUT_WAIT : INT := 6;
END_VAR

(* EDGE DETECTION FOR ALL SENSORS AND SIGNALS *)
SensorFeedEdge := SensorFeed AND NOT PreviousSensorFeed;
SensorWashEdge := SensorWash AND NOT PreviousSensorWash;
SensorWeightEdge := SensorWeight AND NOT PreviousSensorWeight;
SensorFiringEdge := SensorFiring AND NOT PreviousSensorFiring;
SensorOutputEdge := SensorOutput AND NOT PreviousSensorOutput;
WashCompleteEdge := washComplete AND NOT PreviousWashComplete;
WeightCompleteEdge := weightComplete AND NOT PreviousWeightComplete;
FiringCompleteEdge := firingComplete AND NOT PreviousFiringComplete;

(* Update Previous States *)
PreviousSensorFeed := SensorFeed;
PreviousSensorWash := SensorWash;
PreviousSensorWeight := SensorWeight;
PreviousSensorFiring := SensorFiring;
PreviousSensorOutput := SensorOutput;
PreviousWashComplete := washComplete;
PreviousWeightComplete := weightComplete;
PreviousFiringComplete := firingComplete;

(* MANUAL MODE CONTROL *)
IF Mode = FALSE THEN
    (* Interlock: Forward and Reverse cannot be active simultaneously *)
    MotorForward := ForwardButton AND NOT ReverseButton;
    MotorReverse := ReverseButton AND NOT ForwardButton;

    (* Reset automatic mode outputs *)
    kick := FALSE;
    CompletionLight := FALSE;
    firingTemp := 0.0;

    (* Reset state machine *)
    CurrentState := STATE_IDLE;
END_IF

(* AUTOMATIC MODE CONTROL *)
IF Mode = TRUE THEN
    CASE CurrentState OF

        (* STATE_IDLE: Wait for material at loading station *)
        STATE_IDLE:
            MotorForward := FALSE;
            MotorReverse := FALSE;
            kick := FALSE;
            CompletionLight := FALSE;
            firingTemp := 0.0;

            (* Material detected at loading station *)
            IF SensorFeedEdge THEN
                CurrentState := STATE_FEED_DETECTED;
            END_IF

        (* STATE_FEED_DETECTED: Material detected, start motor to move to cleaning *)
        STATE_FEED_DETECTED:
            MotorForward := TRUE;
            MotorReverse := FALSE;
            kick := FALSE;
            CompletionLight := FALSE;

            (* Material reached cleaning station *)
            IF SensorWashEdge THEN
                MotorForward := FALSE;
                CurrentState := STATE_WASH_WAIT;
            END_IF

        (* STATE_WASH_WAIT: Material at cleaning station, wait for washComplete *)
        STATE_WASH_WAIT:
            MotorForward := FALSE;
            MotorReverse := FALSE;
            kick := FALSE;
            CompletionLight := FALSE;

            (* Cleaning complete, move to weighing *)
            IF WashCompleteEdge THEN
                MotorForward := TRUE;
                CurrentState := STATE_WEIGHING_WAIT;
            END_IF

        (* STATE_WEIGHING_WAIT: Material at weighing station, wait for weightComplete *)
        STATE_WEIGHING_WAIT:
            MotorForward := FALSE;
            MotorReverse := FALSE;
            kick := FALSE;
            CompletionLight := FALSE;

            (* Weighing complete, check weight *)
            IF WeightCompleteEdge THEN
                CurrentState := STATE_WEIGHT_CHECK;
            END_IF

        (* STATE_WEIGHT_CHECK: Evaluate weight and determine qualification *)
        STATE_WEIGHT_CHECK:
            weightValue := weight;

            (* Check if weight is within qualified range [100, 200] *)
            IF (weightValue >= 100.0) AND (weightValue <= 200.0) THEN
                (* Qualified product - Calculate firing temperature *)
                (* Linear mapping: weight 100→200 maps to temperature 500→550 *)
                tempCalc := 500.0 + ((weightValue - 100.0) / 100.0) * 50.0;
                firingTemp := tempCalc;
                kick := FALSE;

                (* Move to firing station *)
                MotorForward := TRUE;
                MotorReverse := FALSE;
                CurrentState := STATE_FIRING_WAIT;
            ELSE
                (* Unqualified product - Reject *)
                kick := TRUE;
                firingTemp := 0.0;
                MotorForward := FALSE;
                MotorReverse := FALSE;

                (* Return to idle after rejection *)
                CurrentState := STATE_IDLE;
            END_IF

        (* STATE_FIRING_WAIT: Product at firing station, wait for firingComplete *)
        STATE_FIRING_WAIT:
            kick := FALSE;
            CompletionLight := FALSE;

            (* Firing complete, move to finished product station *)
            IF FiringCompleteEdge THEN
                MotorForward := TRUE;
                MotorReverse := FALSE;
                CurrentState := STATE_OUTPUT_WAIT;
            END_IF

        (* STATE_OUTPUT_WAIT: Product at finished product station *)
        STATE_OUTPUT_WAIT:
            MotorForward := FALSE;
            MotorReverse := FALSE;
            kick := FALSE;

            (* Product detected at output - Turn on completion light *)
            IF SensorOutput THEN
                CompletionLight := TRUE;
            ELSE
                (* Product taken away - Turn off completion light *)
                CompletionLight := FALSE;
                CurrentState := STATE_IDLE;
            END_IF

    END_CASE
END_IF

END_PROGRAM

(* ---- public-medium-03.candidate_02.st ---- *)
{"cmd":["Set-Content -Path 'fb_moving_average.st' -Value @'\nFUNCTION_BLOCK FB_MovingAverage\nVAR_INPUT\n    cyclicExecution : BOOL;\n    trigger : BOOL;\n    value : LREAL;\n    windowSize : INT;\n    reset : BOOL;\nEND_VAR\n\nVAR_OUTPUT\n    average : LREAL;\n    windowSizeReached : BOOL;\n    error : BOOL;\n    status : WORD;\nEND_VAR\n\nVAR\n    buffer : ARRAY[1..100] OF LREAL;\n    index : INT := 1;\n    count : INT := 0;\n    sum : LREAL := 0.0;\n    lastTrigger : BOOL := FALSE;\n    i : INT;\nEND_VAR\n\n(* Main logic *)\nIF reset THEN\n    (* Reset all internal state *)\n    index := 1;\n    count := 0;\n    sum := 0.0;\n    average := 0.0;\n    windowSizeReached := FALSE;\n    error := FALSE;\n    status := 16#0000;\n    \n    (* Clear the buffer *)\n    FOR i := 1 TO 100 DO\n        buffer[i] := 0.0;\n    END_FOR;\n    \n    lastTrigger := FALSE;\n    \nELSIF windowSize < 1 OR windowSize > 100 THEN\n    (* Window size validation error *)\n    error := TRUE;\n    status := 16#8200;\n    windowSizeReached := FALSE;\n    \nELSE\n    (* Check for update condition: cyclic execution OR rising edge of trigger *)\n    IF cyclicExecution OR (trigger AND NOT lastTrigger) THEN\n        (* If buffer is full, subtract the oldest value from sum *)\n        (* If buffer not full, just increment count *)\n        IF count >= windowSize THEN\n            sum := sum - buffer[index];\n        ELSE\n            count := count + 1;\n        END_IF;\n        \n        (* Store new value and update sum *)\n        buffer[index] := value;\n        sum := sum + value;\n        \n        (* Calculate average *)\n        average := sum / LREAL_TO_INT(count);\n        \n        (* Update circular buffer index (wrap around) *)\n        index := (index MOD windowSize) + 1;\n        \n        (* Update windowSizeReached flag *)\n        windowSizeReached := (count >= windowSize);\n        \n        (* Clear error status on successful execution *)\n        error := FALSE;\n        status := 16#0000;\n    END_IF;\n    \n    (* Store trigger state for next cycle (rising edge detection) *)\n    lastTrigger := trigger;\nEND_IF;\n\nEND_FUNCTION_BLOCK\n'@"]}
<newline>
</newline>

{"cmd":["Get-Content -Path 'fb_moving_average.st'"]}
<newline>
</newline>

代码已修复，将 `{ }` 注释语法替换为 ST 标准 `(* *)` 注释语法。

**关键修复：**
- 将所有 `{...}` 注释改为 `(*...*)` 格式
- 保持原有逻辑不变：
  - 循环缓冲区管理（index 从 1 到 windowSize 循环）
  - 上升沿检测（lastTrigger）
  - 窗口大小验证（1-100）
  - 复位功能
  - 状态码（16#0000 成功，16#8200 错误）

(* ---- public-medium-05.candidate_01.st ---- *)
(* Automated Production Line Control *)
(* Three workstations (A→B→C) with manual/automatic mode *)

(* Variable Declarations *)
VAR
    (* Inputs *)
    Mode            : BOOL;  (* 0=Manual, 1=Automatic *)
    ForwardButton   : BOOL;
    ReverseButton   : BOOL;
    SensorA         : BOOL;
    SensorB         : BOOL;
    SensorC         : BOOL;
    ButtonA         : BOOL;
    ButtonB         : BOOL;
    ButtonC         : BOOL;

    (* Outputs *)
    MotorForward    : BOOL;
    MotorReverse    : BOOL;
    CompletionLight : BOOL;

    (* Internal Variables *)
    State           : INT;
END_VAR

(* State Definitions *)
(* 0: IDLE            - Initial/reset state *)
(* 1: AT_STATION_A    - Product at A, waiting for button *)
(* 2: MOVING_TO_B     - Motor moving product from A to B *)
(* 3: AT_STATION_B    - Product at B, waiting for button *)
(* 4: MOVING_TO_C     - Motor moving product from B to C *)
(* 5: AT_STATION_C    - Product at C, waiting for button *)
(* 6: COMPLETE        - Processing complete, light on *)

(* Initialize outputs to OFF *)
MotorForward    := FALSE;
MotorReverse    := FALSE;
CompletionLight := FALSE;

(* MODE SELECTION *)
IF Mode = FALSE THEN
    (* MANUAL MODE *)
    (* Forward and reverse are interlocked - cannot run simultaneously *)
    IF ForwardButton AND NOT ReverseButton THEN
        MotorForward := TRUE;
        MotorReverse := FALSE;
    ELSIF ReverseButton AND NOT ForwardButton THEN
        MotorForward := FALSE;
        MotorReverse := TRUE;
    ELSE
        MotorForward := FALSE;
        MotorReverse := FALSE;
    END_IF

    (* Reset state machine when switching to manual *)
    State := 0;

ELSE
    (* AUTOMATIC MODE *)
    (* State Machine *)
    CASE State OF

        0: (* IDLE - Waiting for product at Station A *)
            MotorForward := FALSE;
            MotorReverse := FALSE;

            IF SensorA THEN
                State := 1;  (* Product arrived at A *)
            END_IF

        1: (* AT STATION A - Waiting for ButtonA *)
            MotorForward := FALSE;
            MotorReverse := FALSE;

            IF ButtonA THEN
                State := 2;  (* Start moving to B *)
            END_IF

        2: (* MOVING TO B - Motor forward *)
            MotorForward := TRUE;
            MotorReverse := FALSE;

            (* Stop when product reaches B *)
            IF SensorB THEN
                MotorForward := FALSE;
                State := 3;
            END_IF

        3: (* AT STATION B - Waiting for ButtonB *)
            MotorForward := FALSE;
            MotorReverse := FALSE;

            IF ButtonB THEN
                State := 4;  (* Start moving to C *)
            END_IF

        4: (* MOVING TO C - Motor forward *)
            MotorForward := TRUE;
            MotorReverse := FALSE;

            (* Stop when product reaches C *)
            IF SensorC THEN
                MotorForward := FALSE;
                State := 5;
            END_IF

        5: (* AT STATION C - Waiting for ButtonC *)
            MotorForward := FALSE;
            MotorReverse := FALSE;

            IF ButtonC THEN
                CompletionLight := TRUE;
                State := 6;  (* Process complete *)
            END_IF

        6: (* COMPLETE - Light on until product removed *)
            MotorForward := FALSE;
            MotorReverse := FALSE;
            CompletionLight := TRUE;

            (* Turn off light when product is taken away *)
            IF NOT SensorC THEN
                CompletionLight := FALSE;
                State := 0;  (* Return to idle for next product *)
            END_IF

    END_CASE
END_IF

(* ---- public-medium-05.candidate_02.st ---- *)
(* Automated Production Line Control *)
(* Three workstations (A→B→C) with manual/automatic mode *)
PROGRAM AutomatedProductionLine
VAR
    (* Inputs *)
    Mode            : BOOL;  (* 0=Manual, 1=Automatic *)
    ForwardButton   : BOOL;
    ReverseButton   : BOOL;
    SensorA         : BOOL;
    SensorB         : BOOL;
    SensorC         : BOOL;
    ButtonA         : BOOL;
    ButtonB         : BOOL;
    ButtonC         : BOOL;

    (* Outputs *)
    MotorForward    : BOOL;
    MotorReverse    : BOOL;
    CompletionLight : BOOL;

    (* Internal Variables *)
    State           : INT;
END_VAR

(* State Definitions *)
(* 0: IDLE            - Initial/reset state *)
(* 1: AT_STATION_A    - Product at A, waiting for button *)
(* 2: MOVING_TO_B     - Motor moving product from A to B *)
(* 3: AT_STATION_B    - Product at B, waiting for button *)
(* 4: MOVING_TO_C     - Motor moving product from B to C *)
(* 5: AT_STATION_C    - Product at C, waiting for button *)
(* 6: COMPLETE        - Processing complete, light on *)

(* Initialize outputs to OFF *)
MotorForward    := FALSE;
MotorReverse    := FALSE;
CompletionLight := FALSE;

(* MODE SELECTION *)
IF Mode = FALSE THEN
    (* MANUAL MODE *)
    (* Forward and reverse are interlocked - cannot run simultaneously *)
    IF ForwardButton AND NOT ReverseButton THEN
        MotorForward := TRUE;
        MotorReverse := FALSE;
    ELSIF ReverseButton AND NOT ForwardButton THEN
        MotorForward := FALSE;
        MotorReverse := TRUE;
    ELSE
        MotorForward := FALSE;
        MotorReverse := FALSE;
    END_IF

    (* Reset state machine when switching to manual *)
    State := 0;

ELSE
    (* AUTOMATIC MODE *)
    (* State Machine *)
    CASE State OF

        0: (* IDLE - Waiting for product at Station A *)
            MotorForward := FALSE;
            MotorReverse := FALSE;

            IF SensorA THEN
                State := 1;  (* Product arrived at A *)
            END_IF

        1: (* AT STATION A - Waiting for ButtonA *)
            MotorForward := FALSE;
            MotorReverse := FALSE;

            IF ButtonA THEN
                State := 2;  (* Start moving to B *)
            END_IF

        2: (* MOVING TO B - Motor forward *)
            MotorForward := TRUE;
            MotorReverse := FALSE;

            (* Stop when product reaches B *)
            IF SensorB THEN
                MotorForward := FALSE;
                State := 3;
            END_IF

        3: (* AT STATION B - Waiting for ButtonB *)
            MotorForward := FALSE;
            MotorReverse := FALSE;

            IF ButtonB THEN
                State := 4;  (* Start moving to C *)
            END_IF

        4: (* MOVING TO C - Motor forward *)
            MotorForward := TRUE;
            MotorReverse := FALSE;

            (* Stop when product reaches C *)
            IF SensorC THEN
                MotorForward := FALSE;
                State := 5;
            END_IF

        5: (* AT STATION C - Waiting for ButtonC *)
            MotorForward := FALSE;
            MotorReverse := FALSE;

            IF ButtonC THEN
                CompletionLight := TRUE;
                State := 6;  (* Process complete *)
            END_IF

        6: (* COMPLETE - Light on until product removed *)
            MotorForward := FALSE;
            MotorReverse := FALSE;
            CompletionLight := TRUE;

            (* Turn off light when product is taken away *)
            IF NOT SensorC THEN
                CompletionLight := FALSE;
                State := 0;  (* Return to idle for next product *)
            END_IF

    END_CASE
END_IF

END_PROGRAM

(* ---- public-medium-06.candidate_01.st ---- *)
(* Slab Thickness Alarm and Fault History Monitor
 * Requirements:
 * 1. Alarm with 500ms minimum hold, active while fault persists
 * 2. Fault counter and 5-entry history (shift register, newest at index 0)
 * 3. Runtime accumulation during normal cutting (valid signal, no fault)
 * 4. Clear state when signal invalid or at power-up
 * 5. Statistics/history are read-only to external callers
 *)
PROGRAM SlabThicknessMonitor
VAR
    (* === Inputs === *)
    THICKNESS_FAULT        : BOOL;   (* Thickness deviation exceeds tolerance *)
    THICKNESS_SIGNAL_VALID : BOOL;   (* Thickness signal validity *)
    CUTTING_RUN            : BOOL;   (* Cutting equipment running status *)
    FaultTimestamp         : DINT;   (* Current timestamp in seconds *)
    CycleTime              : TIME;   (* Elapsed interval for this invocation *)

    (* === Outputs === *)
    THICKNESS_ALARM           : BOOL;                    (* Alarm with min 500ms hold *)
    Slab_Fault_Counter        : UINT;                    (* Valid fault occurrence count *)
    Slab_Runtime_Accumulator  : LTIME;                   (* Accumulated normal runtime *)
    Slab_Fault_History        : ARRAY[0..4] OF DINT;     (* 5 recent fault timestamps *)

    (* === Internal State === *)
    AlarmHoldTimer   : TON;     (* Timer for 500ms alarm hold *)
    FaultWasActive   : BOOL;    (* Rising-edge detection for fault signal *)
    PowerUpComplete  : BOOL;    (* Power-up initialization flag *)
    i                : INT;     (* Loop index for history shift *)
END_VAR

(* === Power-Up Initialization === *)
IF NOT PowerUpComplete THEN
    THICKNESS_ALARM            := FALSE;
    Slab_Fault_Counter         := 0;
    Slab_Runtime_Accumulator   := LTIME#0s;

    FOR i := 0 TO 4 DO
        Slab_Fault_History[i] := 0;
    END_FOR

    FaultWasActive  := FALSE;
    PowerUpComplete := TRUE;
END_IF

(* === Clear State When Signal Invalid === *)
IF NOT THICKNESS_SIGNAL_VALID THEN
    THICKNESS_ALARM  := FALSE;
    AlarmHoldTimer(IN := FALSE);
    FaultWasActive   := FALSE;
ELSE
    (* === Alarm Logic: Immediate activation + 500ms hold === *)
    AlarmHoldTimer(IN  := THICKNESS_FAULT,
                   PT  := T#500ms);
    THICKNESS_ALARM := THICKNESS_FAULT OR AlarmHoldTimer.Q;

    (* === Fault History: Rising-edge detection + shift register === *)
    IF THICKNESS_FAULT AND NOT FaultWasActive THEN
        Slab_Fault_Counter         := Slab_Fault_Counter + 1;
        Slab_Fault_History[4]      := Slab_Fault_History[3];
        Slab_Fault_History[3]      := Slab_Fault_History[2];
        Slab_Fault_History[2]      := Slab_Fault_History[1];
        Slab_Fault_History[1]      := Slab_Fault_History[0];
        Slab_Fault_History[0]      := FaultTimestamp;
    END_IF;

    (* Update fault state for next scan *)
    FaultWasActive := THICKNESS_FAULT;

    (* === Runtime Accumulation: Normal cutting only === *)
    IF CUTTING_RUN AND NOT THICKNESS_FAULT THEN
        Slab_Runtime_Accumulator := Slab_Runtime_Accumulator + CycleTime;
    END_IF
END_IF

END_PROGRAM

(* ---- public-medium-07.candidate_01.st ---- *)
PROGRAM HVAC_Control
VAR
    // Inputs
    OCCUPANCY_DETECTED    : BOOL;
    ENERGY_SAVING_MODE    : BOOL;
    HVAC_MODE_SELECTOR    : INT;

    // Outputs
    SUPPLY_FAN_RUN        : BOOL := FALSE;
    TEMP_SETPOINT_ADJUST  : INT := 0;

    // Internal variables
    occupancy_delay_timer : TON;
END_VAR

//====================================================================
// SUPPLY FAN CONTROL - 30 second delay logic
//====================================================================
// Start 30-second delay when:
//   - Occupancy is detected
//   - Night mode (3) is NOT selected
// Stop immediately and reset timing if:
//   - Occupancy is lost
//   - Night mode is selected
//====================================================================
IF OCCUPANCY_DETECTED AND (HVAC_MODE_SELECTOR <> 3) THEN
    // Start timing with 30-second preset
    occupancy_delay_timer(IN := TRUE, PT := T#30S);

    // Enable fan only after delay completes
    IF occupancy_delay_timer.Q THEN
        SUPPLY_FAN_RUN := TRUE;
    ELSE
        SUPPLY_FAN_RUN := FALSE;
    END_IF;
ELSE
    // Conditions lost - stop fan and reset timer
    occupancy_delay_timer(IN := FALSE);
    SUPPLY_FAN_RUN := FALSE;
END_IF;

//====================================================================
// TEMPERATURE SETPOINT ADJUSTMENT
//====================================================================
// Auto mode (0): 0°C when occupied; +3°C (energy saving) or +2°C (standard) when unoccupied
// Comfort mode (1): 0°C when occupied; +1°C when unoccupied
// Economy mode (2): 0°C when occupied; +4°C when unoccupied
// Night mode (3): +4°C regardless of occupancy
//====================================================================
CASE HVAC_MODE_SELECTOR OF
    0: // Auto mode
        IF OCCUPANCY_DETECTED THEN
            TEMP_SETPOINT_ADJUST := 0;
        ELSE
            IF ENERGY_SAVING_MODE THEN
                TEMP_SETPOINT_ADJUST := 3;
            ELSE
                TEMP_SETPOINT_ADJUST := 2;
            END_IF;
        END_IF;

    1: // Comfort mode
        IF OCCUPANCY_DETECTED THEN
            TEMP_SETPOINT_ADJUST := 0;
        ELSE
            TEMP_SETPOINT_ADJUST := 1;
        END_IF;

    2: // Economy mode
        IF OCCUPANCY_DETECTED THEN
            TEMP_SETPOINT_ADJUST := 0;
        ELSE
            TEMP_SETPOINT_ADJUST := 4;
        END_IF;

    3: // Night mode
        TEMP_SETPOINT_ADJUST := 4;

    ELSE
        TEMP_SETPOINT_ADJUST := 0;
END_CASE;

//====================================================================
// CLAMP TO VALID RANGE ±4°C
//====================================================================
IF TEMP_SETPOINT_ADJUST > 4 THEN
    TEMP_SETPOINT_ADJUST := 4;
ELSIF TEMP_SETPOINT_ADJUST < -4 THEN
    TEMP_SETPOINT_ADJUST := -4;
END_IF;

END_PROGRAM
